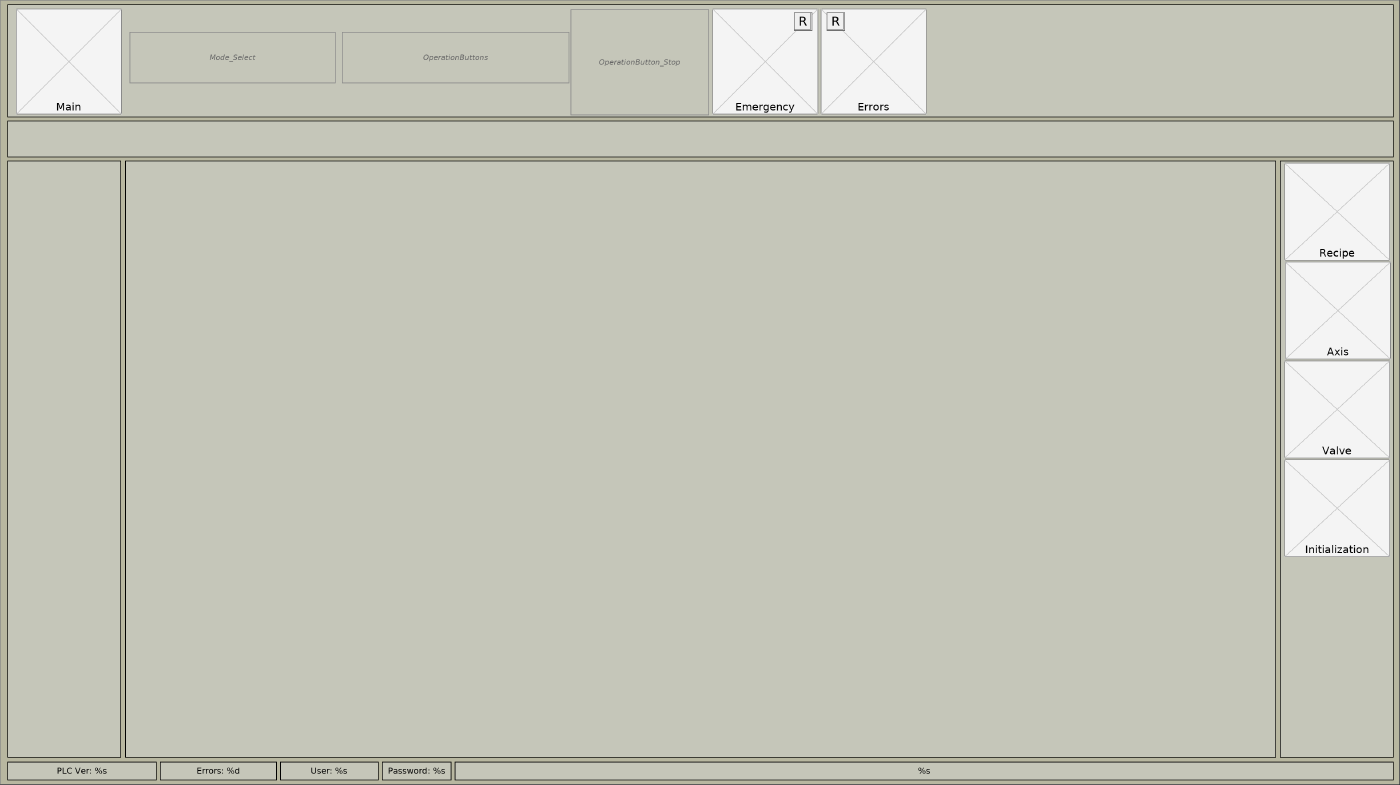
VISUALIZATION TEMP16_9_00_1  // 1924x1080
    Rectangle (0,0 1924x1080)
    Rectangle (385,1048 135x25), "User: %s", text variable: prg_User.actUser
    Rectangle (525,1048 95x25), "Password: %s", text variable: prg_User.Password
        OnMouseDown: write the text variable via Default, min 1, max 999
    Rectangle (220,1048 160x25), "Errors: %d", text variable: Global_Persistent.Errors, colour toggle: Global_Persistent.Errors<>0
        OnMouseUp: execute { Global_Persistent.Errors:=(0); }
    Rectangle (10,1048 205x25), "PLC Ver: %s", text variable: ProgramVersion
    Rectangle (625,1048 1290x25), "%s", text variable: sDateTime
    Rectangle (10,6 1905x155)
    Rectangle (10,166 1905x50)
    Image (22,12 145x145), "Main", image: ImagePool.Main
        OnMouseClick: change screen: vis_MAIN
    Image (979,12 145x145), "Emergency", image: ImagePool.EStop_OK2
        p84334746: GVL_Safety.sBitmap_ESButton
        OnMouseClick: change screen: ES_INT_OPER_16_9
    Image (1128,12 145x145), "Errors", image: ImagePool.Error_No
        p84334746: s_Error_BitmapID
        OnMouseClick: change screen: ERRORS_OPER_16_9
    Button (1136,17 25x25), "R", pressed state: prg_Messages.ResetErrors
        toggle prg_Messages.ResetErrors
    Button (1091,17 25x25), "R"
    Rectangle (10,221 156x821)
    Rectangle (1759,221 156x821)
    Image (1765,224 145x134), "Recipe", image: ImagePool.recipe icon
        OnMouseClick: change screen: Recipe_16_9
    Image (1765,496 145x134), "Valve", image: ImagePool.festo-pistonjpg
        OnMouseClick: change screen: PISTON_OPER_16_9
    Frame (470,44 312x70)
        shows OperationButtons(stOperation := stOpMain)
    Frame (178,44 283x70)
        shows Mode_Select(stMode := stModeMain)
    Image (1765,632 145x134), "Initialization", image: ImagePool.illustration-project-icon
        OnMouseClick: change screen: INIT_OPER_16_9
    Rectangle (172,221 1581x821)
    Frame (784,13 190x145)
        shows OperationButton_Stop(stOperation := stOpMain)
    Image (1766,360 145x134), "Axis", image: ImagePool.ervo-motor-beckhoff
        OnMouseClick: change screen: AXIS_OPER
END_VISUALIZATION

(* stored: Version 1.1.0.1, ProductVersion 3.1.4024.13
   Visu TEMP16_9_00_1: Id {e6a6ea60-81fe-4553-b9fe-912821393375} *)
